(* IEC 61131-3 sources: trust-platform/examples/control/02-derivative-action-and-dynamic-response/32-proportional-position-stiffness/src, 2 files *)

(* ---- Main.st ---- *)
USING Control;

FUNCTION SamePidParameters : BOOL
VAR_INPUT
    Left : Control.PIDParameters;
    Right : Control.PIDParameters;
END_VAR
SamePidParameters :=
    Left.ProportionalGain = Right.ProportionalGain
    AND Left.IntegralGain = Right.IntegralGain
    AND Left.DerivativeGain = Right.DerivativeGain
    AND Left.ProportionalSetpointWeight = Right.ProportionalSetpointWeight
    AND Left.DerivativeSetpointWeight = Right.DerivativeSetpointWeight
    AND Left.Bias = Right.Bias
    AND Left.OutputMinimum = Right.OutputMinimum
    AND Left.OutputMaximum = Right.OutputMaximum
    AND Left.RateMinimum = Right.RateMinimum
    AND Left.RateMaximum = Right.RateMaximum
    AND Left.TrackingTime = Right.TrackingTime
    AND Left.AntiWindup = Right.AntiWindup;
END_FUNCTION

PROGRAM Main
VAR
    Controller : Control.PID;
    (* P position control: Control.PID with zero integral and derivative gains. The output is motor
       torque in N·m, limited to the drive's ±20 N·m. Tune replaces this record. *)
    Parameters : Control.PIDParameters := (
        ProportionalGain := LREAL#4.0,
        IntegralGain := LREAL#0.0,
        DerivativeGain := LREAL#0.0,
        ProportionalSetpointWeight := LREAL#1.0,
        DerivativeSetpointWeight := LREAL#0.0,
        Bias := LREAL#0.0,
        OutputMinimum := LREAL#-20.0,
        OutputMaximum := LREAL#20.0,
        RateMinimum := LREAL#-10000.0,
        RateMaximum := LREAL#10000.0,
        TrackingTime := LREAL#1.0,
        AntiWindup := PIDAntiWindup#BackCalculation
    );
    ConfiguredParameters : Control.PIDParameters;
    ParameterRevision : DINT := 0;
    InitialState : Control.PIDInitialState;
    Input : Control.PIDInput;
    Initialized : BOOL := FALSE;
    AutoMode : BOOL := FALSE;
    ManualTorqueNm : LREAL := 0.0;
    SafetyAbort : BOOL := FALSE;
    SetpointRad : LREAL := 0.0;
    AngleRad : LREAL := 0.0;
    VelocityRadS : LREAL := 0.0;
    TorqueNm : LREAL := 0.0;
    (* Software travel and speed limits of the axis. *)
    AngleLimitRad : LREAL := 2.0;
    VelocityLimitRadS : LREAL := 10.0;
    (* Arrival: the measured velocity at the first sample that reaches a new target. *)
    ArrivalSetpointRad : LREAL := 0.0;
    ApproachRad : LREAL := 0.0;
    Arrived : BOOL := TRUE;
    ArrivalVelocityRadS : LREAL := 0.0;
END_VAR

(* Leaving the travel or speed range removes the torque until a full restart. *)
IF ABS(AngleRad) > AngleLimitRad OR ABS(VelocityRadS) > VelocityLimitRadS THEN
    SafetyAbort := TRUE;
END_IF;

(* Control Studio's Apply replaces this complete record at the task boundary. *)
IF NOT Initialized OR NOT SamePidParameters(Left := Parameters, Right := ConfiguredParameters) THEN
    ConfiguredParameters := Parameters;
    ParameterRevision := ParameterRevision + 1;
END_IF;
Controller.Configure(Parameters := Parameters);

IF NOT Initialized THEN
    (* Hot reset: the axis rests without torque and the setpoint follows the measured angle. *)
    ManualTorqueNm := LREAL#0.0;
    IF NOT AutoMode THEN
        SetpointRad := AngleRad;
    END_IF;
    InitialState.Setpoint := SetpointRad;
    InitialState.ProcessValue := AngleRad;
    InitialState.NominalOutput := ManualTorqueNm;
    InitialState.SaturatedOutput := ManualTorqueNm;
    InitialState.SetpointRate := LREAL#0.0;
    InitialState.ProcessValueRate := LREAL#0.0;
    InitialState.FeedForward := LREAL#0.0;
    Controller.Initialize(State := InitialState);
    ArrivalSetpointRad := SetpointRad;
    Initialized := TRUE;
END_IF;

Input.Setpoint := SetpointRad;
Input.ProcessValue := AngleRad;
Input.CycleTime := LREAL#0.02;
Input.FeedForward := LREAL#0.0;
Input.TrackingOutput := ManualTorqueNm;
IF SafetyAbort THEN
    Input.Mode := PIDMode#Manual;
    Input.ManualOutput := LREAL#0.0;
ELSIF AutoMode AND Parameters.ProportionalGain > LREAL#0.0 THEN
    Input.Mode := PIDMode#Auto;
    Input.ManualOutput := ManualTorqueNm;
ELSE
    Input.Mode := PIDMode#Manual;
    Input.ManualOutput := ManualTorqueNm;
END_IF;
TorqueNm := Controller.Update(Input := Input);

IF SetpointRad <> ArrivalSetpointRad THEN
    ArrivalSetpointRad := SetpointRad;
    ApproachRad := SetpointRad - AngleRad;
    Arrived := FALSE;
END_IF;
IF NOT Arrived AND ApproachRad * (SetpointRad - AngleRad) <= LREAL#0.0 THEN
    Arrived := TRUE;
    ArrivalVelocityRadS := VelocityRadS;
END_IF;

END_PROGRAM

CONFIGURATION Config
RESOURCE Res ON PLC
    TASK MainTask(INTERVAL := T#20ms, PRIORITY := 1);
    PROGRAM P1 WITH MainTask : Main;
END_RESOURCE
VAR_CONFIG
    P1.SafetyAbort AT %MX24.0 : BOOL;
    P1.TorqueNm AT %QL0 : LREAL;
    P1.AngleRad AT %IL0 : LREAL;
    P1.VelocityRadS AT %IL8 : LREAL;
    P1.SetpointRad AT %ML0 : LREAL;
    P1.ManualTorqueNm AT %ML8 : LREAL;
    P1.ArrivalVelocityRadS AT %ML16 : LREAL;
END_VAR
END_CONFIGURATION

(* ---- tests.st ---- *)
(* @trustlsp:runtime-ignore — run these assertions with trust-dev test;
   they are not scheduled PLC instances in the lesson simulator. *)
USING Control;

TEST_PROGRAM TorqueIsProportionalToThePositionError
VAR
    Controller : Control.PID;
    Parameters : Control.PIDParameters;
    Input : Control.PIDInput;
END_VAR
(* The P configuration of Control.PID: Kp = 16 N·m/rad, zero integral and derivative gains. *)
Parameters.ProportionalGain := LREAL#16.0;
Parameters.OutputMinimum := LREAL#-20.0;
Parameters.OutputMaximum := LREAL#20.0;
Parameters.RateMinimum := LREAL#-10000.0;
Parameters.RateMaximum := LREAL#10000.0;
Parameters.TrackingTime := LREAL#1.0;
Controller.Configure(Parameters := Parameters);
Input.Mode := PIDMode#Auto;
Input.CycleTime := LREAL#0.02;
Input.Setpoint := LREAL#1.0;
(* 0.1 rad short of the target: 1.6 N·m. *)
Input.ProcessValue := LREAL#0.9;
ASSERT_NEAR(EXPECTED := LREAL#1.6, ACTUAL := Controller.Update(Input := Input), DELTA := LREAL#1.0e-9);
(* At the target: zero torque, whatever the velocity. *)
Input.ProcessValue := LREAL#1.0;
ASSERT_NEAR(EXPECTED := LREAL#0.0, ACTUAL := Controller.Update(Input := Input), DELTA := LREAL#1.0e-9);
(* 0.2 rad past it: the torque reverses. *)
Input.ProcessValue := LREAL#1.2;
ASSERT_NEAR(EXPECTED := LREAL#-3.2, ACTUAL := Controller.Update(Input := Input), DELTA := LREAL#1.0e-9);
END_TEST_PROGRAM

TEST_PROGRAM TheDriveLimitClipsTheRequest
VAR
    Controller : Control.PID;
    Parameters : Control.PIDParameters;
    Input : Control.PIDInput;
END_VAR
Parameters.ProportionalGain := LREAL#16.0;
Parameters.OutputMinimum := LREAL#-20.0;
Parameters.OutputMaximum := LREAL#20.0;
Parameters.RateMinimum := LREAL#-10000.0;
Parameters.RateMaximum := LREAL#10000.0;
Parameters.TrackingTime := LREAL#1.0;
Controller.Configure(Parameters := Parameters);
Input.Mode := PIDMode#Auto;
Input.CycleTime := LREAL#0.02;
(* A 1.5 rad error requests 24 N·m; the drive delivers at most 20 N·m. *)
Input.Setpoint := LREAL#1.5;
Input.ProcessValue := LREAL#0.0;
ASSERT_NEAR(EXPECTED := LREAL#20.0, ACTUAL := Controller.Update(Input := Input), DELTA := LREAL#1.0e-9);
END_TEST_PROGRAM
